Staubli VAL3: Main.pgx

program Main()
  local bool l_bResult
  local bool l_bStartClock
  local num l_nClock
  local num l_nResult
begin
  //

  home:sVersion="version:5.0"
  resetMotion()
  //初始化
  //  call cycle_Init()
  //
  // userPage("StartUp")

  sMsg=">>> Loading 数据库 "+toString("",saveData:nLibIndex)+" <<<"
  //guohangxin add 2023.03.23
  //call initLib:initlib()
  saveData:nLibIndex=0
  call program:loadPROG(saveData:nLibIndex,l_nResult)
  call trajectory:loadTRAJ(saveData:nLibIndex,l_nResult)
  sMsg=""

  //机器人状态
  taskCreate "plc",60,plc:main()
  wait(taskStatus("plc")==1)
  //HMI
  taskCreate "HMI",50,home:main()
  wait(taskStatus("HMI")==1)
  //  //lifebit
  taskCreate "supervisorTask",10,_supervisorTasks()
  wait(taskStatus("supervisorTask")==1)
  do
    //机器人当前状态
    call _systemStates()
    //生产控制
    call _tCycleCtrl()
    //上下电位置记录
    // call _TolleranceCheck(bAutoConnectMove)
    delay(0)
  until rs:bQuitApp==true

  call kill()

end
